FUNCTION VC_GetUInt16 : UINT
// Reads UInt16 (2 byte, little-endian) from Buf[Pos] and advances Pos.
VAR_IN_OUT
    Buf   : ARRAY[*] OF BYTE;
    Pos   : UDINT;
END_VAR
VAR
    nVal : UINT;
END_VAR

nVal := 0;
VC_GetRaw(Buf := Buf, Pos := Pos, pDst := ADR(nVal), Size := 2);
VC_GetUInt16 := nVal;

END_FUNCTION

(* stored: Version 1.1.0.1, ProductVersion 3.1.4024.12
   POU VC_GetUInt16: Id {bedb9406-c7b6-44d2-adbf-c69564e58d64}, SpecialFunc None *)
